Fanuc KAREL source: kt00076.KL

-- PROVISIONAL review KL for V770-1; original PC SHA256 13e356a34b618f36e77d6afab73f85f85457eb7c7fa701a82a5078ab7c0c7bc2
-- Incomplete behavior may be omitted. Consult companion uncertainty JSON. Do not deploy.
PROGRAM KT00076
%NOLOCKGROUP
VAR
  R1 : REAL
  R2 : REAL
  OUT : REAL
BEGIN
  -- UNRESOLVED_PC offsets 5-16; opcodes 2E,23
  -- UNRESOLVED_PC offsets 21-32; opcodes 2E,23
  -- UNRESOLVED_PC offsets 37-48; opcodes 2E,23
  -- UNRESOLVED_PC offsets 53-64; opcodes 2E,23
  -- UNRESOLVED_PC offsets 69-88; opcodes 21,21,6B,23
  -- UNRESOLVED_PC offsets 93-97; opcodes 7F
END KT00076
